FUNCTION_BLOCK WpfContext EXTENDS TcoCore.TcoContext
VAR
	_serviceModeActive : BOOL;
	{attribute addProperty Name "<#ATEQ G6 PN#>"}
	_ateq1 : TcoAteqMeasurement.TcoAteqG6Pn_v_3_5_x(THIS^);
END_VAR

METHOD PROTECTED Main
IF _serviceModeActive THEN
	_ateq1.Service();
END_IF
_ateq1(inoData := GVL.Ateq1);
END_METHOD

END_FUNCTION_BLOCK

(* stored: Version 1.1.0.1, ProductVersion 3.1.4024.12
   POU WpfContext: Id {709b0734-c343-4049-95ac-3cd974324b35}, SpecialFunc None
   Method Main: Id {b0a973f4-4a76-4e63-b5c5-67f57600aa25} *)
